SUBAPPLICATION Heben_Senken_TO_QDA_PWM_OPC (* 2 Remote-Kommandos (Heben/Senken, je Subscribe+State-Publish, ODER-verknuepft mit IO-Test wie bei ILOCK_SWITCH_2_QXA_OPC) auf 1 ratiometrisches PWM-Signal (Danfoss PVEA: 25%=Senken, 50%=Neutral, 75%=Heben, Lastteiler-korrigiert) + 1 Freigabe-DO als Klick-Toggle (AX_T_FF_INIT, Default AN, per RPC-Methode aus VT und Dashboard aus-/einschaltbar - Not-Bedienung, z.B. Strassenmodus). Generisch fuer jeden PVEA-Aktor mit 2 physischen Kanaelen (links=PWM, rechts=Freigabe), Bedienung von einem Modul ohne eigenes VT. *)
  (* Standard: 61499-2 *)
  (* Version 1.8, 2026-10-15, Franz Höpfinger, Meisterschulen am Ostbahnhof, Kommentar-Korrektur (Franz: 'INIT Kette ueberall so machen, ein REND ist NICHT NOETIG'): FB-Netzwerk war bereits sequenziell (DO_Toggle.INITO -> PWM_Mux.INIT, kein E_REND_2-FB vorhanden), aber der INITO-Comment beschrieb noch faelschlich ein Rendezvous aus der v1.7-Planung. Nur Dokumentation angepasst, keine funktionale Aenderung. *)
  (* Version 1.7, 2026-10-13, Franz Höpfinger, Meisterschulen am Ostbahnhof, Neuer SubAppEventOutput INITO (Type EInit) fuer Aufnahme_Option.SUB (Option::AOption-Socket-Wrapper, analog Bunker_Klappen_Option.SUB) - PWM_Mux.INITO (HebenSenken_ILOCK_QDA_PWM_OPC v1.6) UND DO_Toggle.INITO (DO_TOGGLE_RPC_QXA_OPC v1.3) sind 2 echte, unabhaengige physische Kanal-Confirms (PWM-Kanal + Freigabe-DO-Kanal). E_REND_2 (Rendezvous/AND, nicht E_MERGE_2/OR) wartet auf BEIDE bevor INITO genau 1x feuert - ein nachgelagerter AOption-Socket (DEMUX Break-before-Make) erwartet pro Umschaltvorgang genau 1 INIT_CNF, ein doppeltes Feuern waere dort undefiniert. INIT selbst resettet E_REND_2 (R), damit jeder neue INIT-Zyklus wieder auf beide wartet. *)
  (* Version 1.6, 2026-10-11, Franz Höpfinger, Meisterschulen am Ostbahnhof, Neuer SubAppEventInput INIT (Type EInit), durchgereicht an PWM_Mux.INIT (HebenSenken_ILOCK_QDA_PWM_OPC v1.5) UND DO_Toggle.INIT (DO_TOGGLE_RPC_QXA_OPC v1.2) statt Auto-Verteilung - analog ILOCK_SWITCH_2_QXA_OPC v1.2, 'Init wie bei Tecu' (Franz). *)
  (* Version 1.5, 2026-10-11, Franz Höpfinger, Meisterschulen am Ostbahnhof, Neuer QI-InputVar (Default TRUE, rueckwaertskompatibel) durchgereicht an PWM_Mux.QI (HebenSenken_ILOCK_QDA_PWM_OPC v1.4) UND DO_Toggle.QI (DO_TOGGLE_RPC_QXA_OPC v1.1) - analog ILOCK_SWITCH_2_QXA_OPC v1.1, haelt beide physischen Kanaele dieser Instanz gemeinsam inaktiv. *)
  (* Version 1.4, 2026-09-20, Franz Höpfinger, Meisterschulen am Ostbahnhof, PWM_POW-Socket ergaenzt (reiner Passthrough an PWM_Mux.PWM_POW), da HebenSenken_ILOCK_QDA_PWM_OPC v1.1 PWM_POW jetzt als eigenen Socket statt intern fest 1.0 hat - jeder Aufrufer muss ihn jetzt verbinden. *)
  (* Version 1.3, 2026-09-08, Franz Höpfinger, Meisterschulen am Ostbahnhof, V1.1: IO-Test fuer Heben/Senken ergaenzt (SUBSCRIBE_TEST_HEBEN/SENKEN, ODER vor dem ILOCK), Publish-Punkte (State+Test) hinter den ILOCK verlegt (wie ILOCK_SWITCH_2_QXA_OPC), Freigabe-DO von starrem initval_AX auf AX_T_FF_INIT-Klick-Toggle per RPC-Methode umgestellt - KEIN OR nach dem Flipflop, AX_T_FF_INIT.Q ist alleinige Source of Truth fuer den Ausgang. V1.2: Freigabe-DO-Teilnetz nach MyLib::sys::DO_TOGGLE_RPC_QXA_OPC ausgelagert. V1.3: PWM/ILOCK/Mux-Teilnetz nach MyLib::sys::HebenSenken_ILOCK_QDA_PWM_OPC ausgelagert - diese SubApp ist jetzt nur noch die Zusammensetzung beider Bausteine, Schnittstelle unveraendert. *)
  PACKAGE MyLib::sys;
  IMPORT logiBUS::io::DQ::logiBUS_DO;
  IMPORT logiBUS::io::DQ::logiBUS_DO_S;
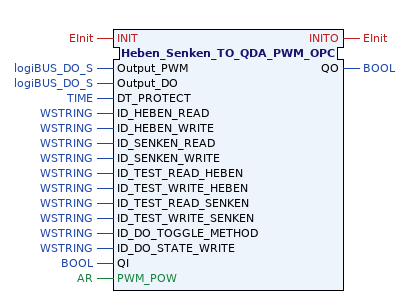
  EVENT_INPUT
    INIT : EInit; (* Initialisierung - vom Aufrufer sequenziert statt per Auto-Verteilung, damit QI vor der physischen Kanalbindung feststeht *)
  END_EVENT
  EVENT_OUTPUT
    INITO : EInit; (* Initialisierung abgeschlossen - sequenzielles Confirm: DO_Toggle zuerst, dann PWM_Mux (kein Rendezvous noetig, beide sind reine physische Ausgangskanaele) *)
  END_EVENT
  VAR_INPUT
    Output_PWM : logiBUS::io::DQ::logiBUS_DO_S := logiBUS_DO::Invalid; (* Physischer PWM-Ausgang (linker Kanal): 25/50/75% Tastgrad, ratiometrisch *)
    Output_DO : logiBUS::io::DQ::logiBUS_DO_S := logiBUS_DO::Invalid; (* Physischer Freigabe-Ausgang (rechter Kanal): Klick-Toggle, Default AN *)
    DT_PROTECT : TIME := T#300ms; (* Schutz-Totzeit vor Richtungswechsel *)
    ID_HEBEN_READ : WSTRING; (* Echtes Funktions-Kommando Heben (Subscribe) *)
    ID_HEBEN_WRITE : WSTRING; (* Echte Funktions-Rueckmeldung Heben, HINTER dem ILOCK (Publish) *)
    ID_SENKEN_READ : WSTRING; (* Echtes Funktions-Kommando Senken (Subscribe) *)
    ID_SENKEN_WRITE : WSTRING; (* Echte Funktions-Rueckmeldung Senken, HINTER dem ILOCK (Publish) *)
    ID_TEST_READ_HEBEN : WSTRING; (* Bestehende IO-Test-Subscribe-Adresse Heben (z.B. STG2_Q0x_READ), ODER-verknuepft mit ID_HEBEN_READ vor dem ILOCK *)
    ID_TEST_WRITE_HEBEN : WSTRING; (* Bestehende IO-Test-Publish-Adresse Heben, HINTER dem ILOCK (z.B. STG2_Q0x_WRITE) *)
    ID_TEST_READ_SENKEN : WSTRING; (* Bestehende IO-Test-Subscribe-Adresse Senken, ODER-verknuepft mit ID_SENKEN_READ vor dem ILOCK *)
    ID_TEST_WRITE_SENKEN : WSTRING; (* Bestehende IO-Test-Publish-Adresse Senken, HINTER dem ILOCK *)
    ID_DO_TOGGLE_METHOD : WSTRING; (* Lokale Methodenadresse (ACTION=CREATE_METHOD) fuer den argumentlosen Freigabe-Toggle-Trigger - wird von STG1 (SoftKey-Relay) UND direkt vom OPC-Dashboard (CALL_METHOD) aufgerufen, beide Aufrufer teilen sich denselben Flipflop-Takt *)
    ID_DO_STATE_WRITE : WSTRING; (* Lokale Publish-Adresse (ACTION=WRITE) fuer den tatsaechlichen Freigabe-Zustand (AX_T_FF_INIT.Q) - wird von VT und Dashboard remote abonniert *)
    QI : BOOL := TRUE; (* Qualifier fuer beide physischen Ausgaenge (PWM+Freigabe-DO) - FALSE haelt diese Instanz komplett inaktiv (keine Hardware-Bindung), fuer den Fall dass derselbe physische Kanal je nach Maschinenvariante anderweitig genutzt wird *)
  END_VAR
  VAR_OUTPUT
    QO : BOOL; (* Quality Output - TRUE if service executed successfully (AND aus PWM_Mux/DO_Toggle) *)
  END_VAR
  SOCKETS
    PWM_POW : adapter::types::unidirectional::AR; (* PWM Power 1.0 = Maximale Power, 0.0 = Aus, 0.5 = Halb - durchgereicht an PWM_Mux.PWM_POW *)
  END_SOCKETS
  FBS
    AND_QO : iec61131::booleanOperators::AND_BOOL_2;
  END_FBS
  SUBAPPS
    PWM_Mux : MyLib::sys::HebenSenken_ILOCK_QDA_PWM_OPC;
    DO_Toggle : MyLib::sys::DO_TOGGLE_RPC_QXA_OPC;
  END_SUBAPPS
  EVENT_CONNECTIONS
    INIT TO DO_Toggle.INIT;
    PWM_Mux.INITO TO INITO;
    PWM_Mux.INITO TO AND_QO.REQ;
    DO_Toggle.INITO TO PWM_Mux.INIT;
  END_CONNECTIONS
  DATA_CONNECTIONS
    ID_HEBEN_READ TO PWM_Mux.ID_HEBEN_READ;
    ID_TEST_READ_HEBEN TO PWM_Mux.ID_TEST_READ_HEBEN;
    ID_TEST_WRITE_HEBEN TO PWM_Mux.ID_TEST_WRITE_HEBEN;
    ID_HEBEN_WRITE TO PWM_Mux.ID_HEBEN_WRITE;
    ID_SENKEN_READ TO PWM_Mux.ID_SENKEN_READ;
    ID_TEST_READ_SENKEN TO PWM_Mux.ID_TEST_READ_SENKEN;
    ID_TEST_WRITE_SENKEN TO PWM_Mux.ID_TEST_WRITE_SENKEN;
    ID_SENKEN_WRITE TO PWM_Mux.ID_SENKEN_WRITE;
    Output_PWM TO PWM_Mux.Output_PWM;
    DT_PROTECT TO PWM_Mux.DT_PROTECT;
    Output_DO TO DO_Toggle.Output_DO;
    ID_DO_TOGGLE_METHOD TO DO_Toggle.ID_DO_TOGGLE_METHOD;
    ID_DO_STATE_WRITE TO DO_Toggle.ID_DO_STATE_WRITE;
    QI TO PWM_Mux.QI;
    QI TO DO_Toggle.QI;
    PWM_Mux.QO TO AND_QO.IN1;
    DO_Toggle.QO TO AND_QO.IN2;
    AND_QO.OUT TO QO;
  END_CONNECTIONS
  ADAPTER_CONNECTIONS
    PWM_POW TO PWM_Mux.PWM_POW;
  END_CONNECTIONS
END_SUBAPPLICATION
